// TIA Portal V14 SP1 export
// export: Created 2000-01-01T00:00:00.0000000Z, ExportSetting None
DATA_BLOCK "MCP_RC_DB2"   // DB9803
{ S7_Optimized_Access := 'FALSE' }
   VAR
      Ready : Bool := FALSE;
   END_VAR
BEGIN
END_DATA_BLOCK
